(* IEC 61131-3 sources: BODAS-HelloWorld/st/bodas_rc18_12_40/plc_logic/application/02_easyconfig/easyconfig_import/bds_in_ec, 7 files *)

(* ---- bds_indig_signal_te-bds_inDig_signal_te.st ---- *)
(* --- Interface --- *)
///BODAS configuration of available digital input signals
{attribute 'qualified_only' := ''}
{attribute 'strict' := ''}
TYPE bds_inDig_signal_te : (
		bds_inDig_K22_E := 0,
		///End V1
		bds_inDig_K21_E,
		bds_inDig_numSignal_E
	) USINT;
END_TYPE

(* ---- bds_ini_signal_te-bds_inI_signal_te.st ---- *)
(* --- Interface --- *)
///BODAS configuration of available current measurement input signals
{attribute 'qualified_only' := ''}
{attribute 'strict' := ''}
TYPE bds_inI_signal_te : (
		bds_inI_A38_E := 0,
		bds_inI_A39_E,
		bds_inI_K37_E,
		bds_inI_K30_E,
		///End V1
		bds_inI_A43_E,
		bds_inI_numSignal_E
	) USINT;
END_TYPE

(* ---- bds_inpha_signal_te-bds_inPha_signal_te.st ---- *)
(* --- Interface --- *)
{attribute 'external_name' := 'cmp_rts_bds_inPha_signal_te'}
TYPE bds_inPha_signal_te : (
		bds_inPha_K55_K61_E := 0,
		bds_inPha_numSignal_E
	) USINT;
END_TYPE

(* ---- bds_inpwm_signal_te-bds_inPwm_signal_te.st ---- *)
(* --- Interface --- *)
///Definition of input signals for PWM
{attribute 'qualified_only' := ''}
{attribute 'strict' := ''}
TYPE bds_inPwm_signal_te : (
		bds_inPwm_K54_E := 0,
		bds_inPwm_K37_E,
		bds_inPwm_K30_E,
		bds_inPwm_A43_E,
		bds_inPwm_A59_A44_E,
		bds_inPwm_numSignal_E
	) USINT;
END_TYPE

(* ---- bds_inr_signal_te-bds_inR_signal_te.st ---- *)
(* --- Interface --- *)
///Definition of input signals for Resistance
{attribute 'qualified_only' := ''}
{attribute 'strict' := ''}
TYPE bds_inR_signal_te : (
		bds_inR_K41_E := 0,
		bds_inR_K65_E,
		bds_inR_K63_E,
		bds_inR_K64_E,
		bds_inR_K32_E,
		bds_inR_K33_E,
		bds_inR_numSignal_E
	) USINT;
END_TYPE

(* ---- bds_inu_signal_te-bds_inU_signal_te.st ---- *)
(* --- Interface --- *)
///Definition of  input Configured Signals for Voltage( Consists signals of all variants)
{attribute 'qualified_only' := ''}
{attribute 'strict' := ''}
TYPE bds_inU_signal_te : (
		bds_inU_K52_E := 0,
		bds_inU_K60_E,
		bds_inU_K43_E,
		bds_inU_K54_E,
		bds_inU_K55_E,
		bds_inU_K39_E,
		bds_inU_K38_E,
		bds_inU_K40_E,
		bds_inU_K42_E,
		bds_inU_K37_E,
		bds_inU_K61_E,
		bds_inU_K45_E,
		bds_inU_K44_E,
		bds_inU_A21_E,
		bds_inU_A36_E,
		bds_inU_A37_E,
		bds_inU_A38_E,
		bds_inU_A39_E,
		bds_inU_K30_E,
		bds_inU_A43_E,
		bds_inU_A22_E,
		bds_inU_A23_E,
		bds_inU_A24_E,
		bds_inU_K78_E,
		bds_inU_K76_E,
		bds_inU_K74_E,
		bds_inU_K77_E,
		bds_inU_K10_E,
		bds_inU_K75_E,
		bds_inU_K31_E,
		bds_inU_K34_E,
		bds_inU_A13_E,
		bds_inU_A40_E,
		bds_inU_A41_E,
		bds_inU_A42_E,
		bds_inU_A25_E,
		bds_inU_A26_E,
		bds_inU_A27_E,
		bds_inU_A14_E,
		bds_inU_A57_E,
		bds_inU_A28_E,
		bds_inU_A29_E,
		bds_inU_K11_E,
		bds_inU_K35_E,
		bds_inU_A59_E,
		bds_inU_numSignal_E
	) USINT;
END_TYPE

(* ---- bds_in_ec_gvl-bds_in_ec_gvl.st ---- *)
(* --- Interface --- *)
{attribute 'qualified_only' := ''}
VAR_GLOBAL CONSTANT
	BDS_inCmn_postVariants_DU8 : USINT := 1;
END_VAR
